(* IEC 61131-3 sources: s7-to-codesys/tests/POUs/S7Compat/FB_F_NormX_Test, 9 files *)

(* ---- FB_F_NormX_Test.decl.st ---- *)
// Назначение: набор тестов CfUnit (coUnit 1.2.0.0) для F_NormX — аналога S7 NORM_X:
//             середина и границы диапазона 0…27648, значения ниже и выше диапазона
//             (линейное продолжение), обратный диапазон (та же формула) и вырожденный
//             диапазон (0.0 — решение s7conv). Ожидаемые значения — по формуле Siemens
//             OUT = (VALUE - MIN) / (MAX - MIN), а не по результату реализации.
//             Экземпляр набора объявляется в PRG_Tests (объявление регистрирует набор).
// Автор:      kr0nsch
// Версия:     0.1.0
// Документ:   docs/MAPPING.md, раздел «NORM_X и SCALE_X»
FUNCTION_BLOCK FB_F_NormX_Test EXTENDS coUnit.FB_TestSuite
VAR CONSTANT
    // арифметика REAL: сравнение с допуском
    R_DELTA : REAL := 0.0001;
END_VAR

(* ---- AboveMaxExtrapolates.method.decl.st ---- *)
// F_NormX(rMin := 0.0, rValue := 30412.8, rMax := 27648.0) = 1.1.
METHOD PRIVATE AboveMaxExtrapolates
VAR
    rResult : REAL;     // результат F_NormX
END_VAR

(* ---- AtMaxGivesOne.method.decl.st ---- *)
// F_NormX(rMin := 0.0, rValue := 27648.0, rMax := 27648.0) = 1.0.
METHOD PRIVATE AtMaxGivesOne
VAR
    rResult : REAL;     // результат F_NormX
END_VAR

(* ---- AtMinGivesZero.method.decl.st ---- *)
// F_NormX(rMin := 0.0, rValue := 0.0, rMax := 27648.0) = 0.0.
METHOD PRIVATE AtMinGivesZero
VAR
    rResult : REAL;     // результат F_NormX
END_VAR

(* ---- BelowMinExtrapolates.method.decl.st ---- *)
// F_NormX(rMin := 0.0, rValue := -2764.8, rMax := 27648.0) = -0.1.
METHOD PRIVATE BelowMinExtrapolates
VAR
    rResult : REAL;     // результат F_NormX
END_VAR

(* ---- EqualBoundsGivesZero.method.decl.st ---- *)
// F_NormX(rMin := 5.0, rValue := 5.0, rMax := 5.0) = 0.0.
METHOD PRIVATE EqualBoundsGivesZero
VAR
    rResult : REAL;     // результат F_NormX
END_VAR

(* ---- MidRangeGivesHalf.method.decl.st ---- *)
// F_NormX(rMin := 0.0, rValue := 13824.0, rMax := 27648.0) = 0.5.
METHOD PRIVATE MidRangeGivesHalf
VAR
    rResult : REAL;     // результат F_NormX
END_VAR

(* ---- OffsetRange.method.decl.st ---- *)
// F_NormX(rMin := 4.0, rValue := 12.0, rMax := 20.0) = 0.5.
METHOD PRIVATE OffsetRange
VAR
    rResult : REAL;     // результат F_NormX
END_VAR

(* ---- ReversedBoundsKeepsFormula.method.decl.st ---- *)
// F_NormX(rMin := 100.0, rValue := 75.0, rMax := 0.0) = 0.25.
METHOD PRIVATE ReversedBoundsKeepsFormula
VAR
    rResult : REAL;     // результат F_NormX
END_VAR
